(* IEC 61131-3 sources: codesys-framework/txt/application/WeVe Core (library)/60 Event/FB_EventGroup/Protected, 2 files *)

(* ---- Configure.method.st ---- *)
// Config van één event invullen. De bron (nSubMachine, nSubMachineId) komt van de groep,
// zodat elke instantie van een module zijn eigen bron heeft met dezelfde event-ID's.
// FALSE bij een ongeldige index.
METHOD PROTECTED Configure : BOOL
VAR_INPUT
	iEvent 			: INT;
	udiEventId 		: UDINT;
	eEventLevel 	: E_EventLevels;
	xResetable 		: BOOL;
	sMessage 		: STRING(GVL_Logger.cMaxMessageLength);		// placeholders %0..%9
END_VAR
VAR
	fbEvent 		: I_Event;
	scConfig 		: SC_Event;
END_VAR

// --- BEGIN IMPLEMENTATION ---

fbEvent := GetEvent(iEvent);

IF fbEvent = 0 THEN
	Configure := FALSE;
	RETURN;
END_IF

scConfig.udiEventId 	:= udiEventId;
scConfig.nSubMachine 	:= _nSubMachine;
scConfig.nSubMachineId 	:= _nSubMachineId;
scConfig.eEventLevel 	:= eEventLevel;
scConfig.xResetable 	:= xResetable;
scConfig.sMessage 		:= sMessage;

fbEvent.Config := scConfig;
Configure := TRUE;

(* ---- ConfigureEvents.method.st ---- *)
// Door de afgeleide groep: één Configure-regel per event. Wordt aangeroepen vanuit Initialize.
//   Configure(E_AirPressureEvent.PressureNok, cEv_MainPressureNotOk, E_EventLevels.EventIsAlarm_SupervisorLevel, TRUE,  'Invalid air pressure');
//   Configure(E_AirPressureEvent.PressureLow, cEv_MainPressureLow,   E_EventLevels.EventIsWarning_Urgent,        FALSE, 'Air pressure low: %0 bar');
METHOD PROTECTED ABSTRACT ConfigureEvents
VAR_INPUT
END_VAR
